// TIA Portal V21 export
// export: Created 2026-11-21T13:31:41.3155978Z, ExportSetting WithDefaults, DisplayName Totally Integrated Automation Portal, DisplayVersion V21, DisplayName STEP 7 Professional, DisplayVersion V21, DisplayName STEP 7 Safety, DisplayVersion V21, DisplayName Tech WebApplication, DisplayVersion V21, DisplayName WinCC Basic/Comfort/Advanced, DisplayVersion V21, DisplayName WinCC Unified, DisplayVersion V21
FUNCTION_BLOCK "ClassicFbd"   // FB11, FBD
TITLE = ClassicFbd
VERSION : 0.1
// Function block diagram on a classic CPU.
// stored: AutoNumber true, IsIECCheckEnabled false, UDAEnableTagReadback false
   VAR_INPUT
      enable : Bool;
   END_VAR
   VAR_OUTPUT
      running : Bool;
   END_VAR
   VAR DB_SPECIFIC
      latched : Bool;
   END_VAR
BEGIN

REGION Network 1: Latch
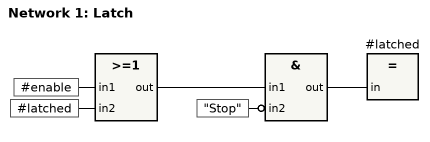
   #latched := (#enable OR #latched) AND NOT "Stop";
END_REGION
END_FUNCTION_BLOCK
